FUNCTION_BLOCK fbMonoSwitch IMPLEMENTS iSwitch
VAR_INPUT
	Input AT %I* : BOOL;
END_VAR					// Physical switch input
VAR
	RTrigInput : R_TRIG;
	FTrigInput : F_TRIG;
END_VAR

RTrigInput(CLK := Input);
FTrigInput(CLK := Input);

PROPERTY IsPressed : BOOL
GET
IsPressed := THIS^.Input;
END_GET
END_PROPERTY

PROPERTY IsReleased : BOOL
GET
IsReleased := NOT THIS^.Input;
END_GET
END_PROPERTY

PROPERTY PUBLIC OnPressed : BOOL
GET
OnPressed := RTrigInput.Q;
END_GET
END_PROPERTY

PROPERTY OnReleased : BOOL
GET
OnReleased := FTrigInput.Q;
END_GET
END_PROPERTY

END_FUNCTION_BLOCK

(* stored: Version 1.1.0.1
   POU fbMonoSwitch: Id {21737aef-df48-4987-83e0-aae9b7cbc7ab}, SpecialFunc None
   Property IsPressed: Id {3ddc41e3-a43a-457c-8835-114dca2b3407}
   Get Get: Id {61dbcbff-306a-4c29-b7b4-947c3ee82b24}
   Property IsReleased: Id {6c0ebfae-fd6b-467c-bcf0-d0f0949b6be2}
   Get Get: Id {1b38215a-e5dc-40a6-900f-84342805f4f2}
   Property OnPressed: Id {238fedb4-7f31-449e-bffb-88405f0e3fe6}
   Get Get: Id {bc4b2b4d-b425-4031-ada5-782516be3c69}
   Property OnReleased: Id {f2e12f74-1423-4b11-9d68-63053027c6bb}
   Get Get: Id {00b0c95b-d4ed-4500-978f-f246b06ade20} *)
